SYSTEM PID_Identification_Observer (* Synthetic observation only; native export and execution pending *)
  APPLICATION Observer_Test (* Fixed PID; no gain-update connections *)
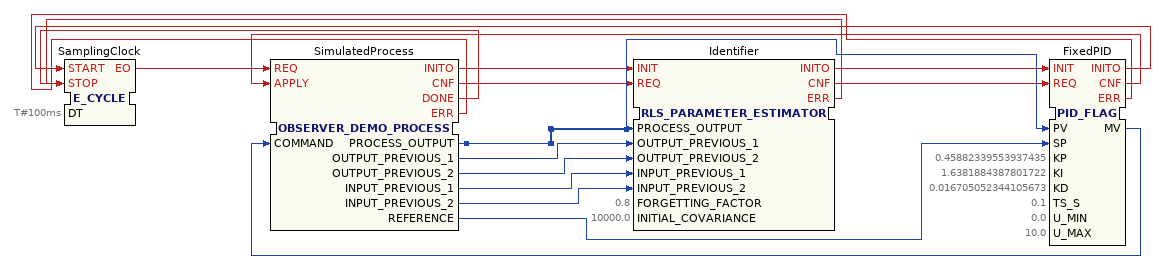
    FBS
      SamplingClock : E_CYCLE(DT := T#100ms);
      SimulatedProcess : OBSERVER_DEMO_PROCESS;
      Identifier : RLS_PARAMETER_ESTIMATOR(FORGETTING_FACTOR := 0.8, INITIAL_COVARIANCE := 10000.0);
      FixedPID : PID_FLAG(KP := 0.45882339553937435, KI := 1.6381884387801722, KD := 0.016705052344105673, TS_S := 0.1, U_MIN := 0.0, U_MAX := 10.0);
    END_FBS
    EVENT_CONNECTIONS
      SimulatedProcess.INITO TO Identifier.INIT;
      Identifier.INITO TO FixedPID.INIT;
      FixedPID.INITO TO SamplingClock.START;
      SamplingClock.EO TO SimulatedProcess.REQ;
      SimulatedProcess.CNF TO Identifier.REQ;
      Identifier.CNF TO FixedPID.REQ;
      FixedPID.CNF TO SimulatedProcess.APPLY;
      SimulatedProcess.DONE TO SamplingClock.STOP;
      SimulatedProcess.ERR TO SamplingClock.STOP;
      Identifier.ERR TO SamplingClock.STOP;
      FixedPID.ERR TO SamplingClock.STOP;
    END_CONNECTIONS
    DATA_CONNECTIONS
      SimulatedProcess.PROCESS_OUTPUT TO Identifier.PROCESS_OUTPUT;
      SimulatedProcess.OUTPUT_PREVIOUS_1 TO Identifier.OUTPUT_PREVIOUS_1;
      SimulatedProcess.OUTPUT_PREVIOUS_2 TO Identifier.OUTPUT_PREVIOUS_2;
      SimulatedProcess.INPUT_PREVIOUS_1 TO Identifier.INPUT_PREVIOUS_1;
      SimulatedProcess.INPUT_PREVIOUS_2 TO Identifier.INPUT_PREVIOUS_2;
      SimulatedProcess.PROCESS_OUTPUT TO FixedPID.PV;
      SimulatedProcess.REFERENCE TO FixedPID.SP;
      FixedPID.MV TO SimulatedProcess.COMMAND;
    END_CONNECTIONS
  END_APPLICATION
  DEVICE LocalObserver : FORTE_PC(MGR_ID := "localhost:61499") (* Local synthetic test only *)
    {SET_ATTRIBUTE(Profile, HOLOBLOC)}
    RESOURCE EMB_RES : EMB_RES
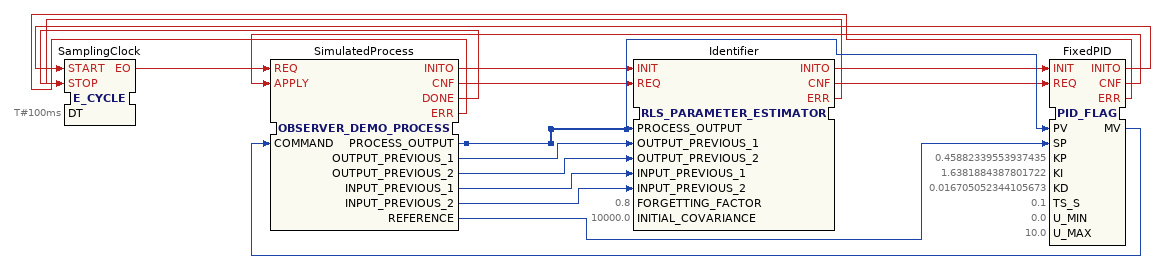
      FBS
        SamplingClock : E_CYCLE(DT := T#100ms);
        SimulatedProcess : OBSERVER_DEMO_PROCESS;
        Identifier : RLS_PARAMETER_ESTIMATOR(FORGETTING_FACTOR := 0.8, INITIAL_COVARIANCE := 10000.0);
        FixedPID : PID_FLAG(KP := 0.45882339553937435, KI := 1.6381884387801722, KD := 0.016705052344105673, TS_S := 0.1, U_MIN := 0.0, U_MAX := 10.0);
      END_FBS
      EVENT_CONNECTIONS
        SimulatedProcess.INITO TO Identifier.INIT;
        Identifier.INITO TO FixedPID.INIT;
        FixedPID.INITO TO SamplingClock.START;
        SamplingClock.EO TO SimulatedProcess.REQ;
        SimulatedProcess.CNF TO Identifier.REQ;
        Identifier.CNF TO FixedPID.REQ;
        FixedPID.CNF TO SimulatedProcess.APPLY;
        SimulatedProcess.DONE TO SamplingClock.STOP;
        SimulatedProcess.ERR TO SamplingClock.STOP;
        Identifier.ERR TO SamplingClock.STOP;
        FixedPID.ERR TO SamplingClock.STOP;
      END_CONNECTIONS
      DATA_CONNECTIONS
        SimulatedProcess.PROCESS_OUTPUT TO Identifier.PROCESS_OUTPUT;
        SimulatedProcess.OUTPUT_PREVIOUS_1 TO Identifier.OUTPUT_PREVIOUS_1;
        SimulatedProcess.OUTPUT_PREVIOUS_2 TO Identifier.OUTPUT_PREVIOUS_2;
        SimulatedProcess.INPUT_PREVIOUS_1 TO Identifier.INPUT_PREVIOUS_1;
        SimulatedProcess.INPUT_PREVIOUS_2 TO Identifier.INPUT_PREVIOUS_2;
        SimulatedProcess.PROCESS_OUTPUT TO FixedPID.PV;
        SimulatedProcess.REFERENCE TO FixedPID.SP;
        FixedPID.MV TO SimulatedProcess.COMMAND;
      END_CONNECTIONS
    END_RESOURCE
  END_DEVICE
  MAPPINGS
    Observer_Test.SamplingClock ON LocalObserver.EMB_RES.SamplingClock;
    Observer_Test.SimulatedProcess ON LocalObserver.EMB_RES.SimulatedProcess;
    Observer_Test.Identifier ON LocalObserver.EMB_RES.Identifier;
    Observer_Test.FixedPID ON LocalObserver.EMB_RES.FixedPID;
  END_MAPPINGS
END_SYSTEM
